(* IEC 61131-3 sources: llm-plc-st-eval/data/processed/gpt-4o/B4/zero_shot, 3 files *)

(* ---- ejec_1.st ---- *)
FUNCTION_BLOCK FB_Giro
VAR_INPUT
    btnFwd : BOOL;   // Botón para giro en sentido horario
    btnRev : BOOL;   // Botón para giro en sentido antihorario
    btnParo : BOOL;  // Botón de paro
END_VAR

VAR_OUTPUT
    fwd : BOOL;      // Salida para giro en sentido horario
    rev : BOOL;      // Salida para giro en sentido antihorario
END_VAR

VAR
    estado : INT;    // Estado actual del motor
END_VAR

// Estados posibles
// 0: Parado
// 1: Girando en sentido horario
// 2: Girando en sentido antihorario

// Lógica de control
IF btnParo THEN
    // Si se presiona el botón de paro, el motor se detiene
    estado := 0;
ELSIF btnFwd AND (estado = 0) THEN
    // Si se presiona el botón de giro horario y el motor está parado
    estado := 1;
ELSIF btnRev AND (estado = 0) THEN
    // Si se presiona el botón de giro antihorario y el motor está parado
    estado := 2;
END_IF

// Actualización de salidas según el estado
CASE estado OF
    0: // Parado
        fwd := FALSE;
        rev := FALSE;
    1: // Girando en sentido horario
        fwd := TRUE;
        rev := FALSE;
    2: // Girando en sentido antihorario
        fwd := FALSE;
        rev := TRUE;
END_CASE

END_FUNCTION_BLOCK

(* ---- ejec_2.st ---- *)
FUNCTION_BLOCK FB_Giro
VAR_INPUT
    btnFwd : BOOL;    // Botón para giro en sentido horario
    btnRev : BOOL;    // Botón para giro en sentido antihorario
    btnParo : BOOL;   // Botón de paro
END_VAR

VAR_OUTPUT
    fwd : BOOL := FALSE;  // Salida para giro en sentido horario
    rev : BOOL := FALSE;  // Salida para giro en sentido antihorario
END_VAR

VAR
    estado : INT := 0;    // Estado del motor: 0 = Parado, 1 = Horario, 2 = Antihorario
END_VAR

// Lógica de control del motor
IF btnParo THEN
    // Si se presiona el botón de paro, detener el motor
    fwd := FALSE;
    rev := FALSE;
    estado := 0;
ELSIF btnFwd AND (estado = 0) THEN
    // Si se presiona el botón de giro horario y el motor está parado
    fwd := TRUE;
    rev := FALSE;
    estado := 1;
ELSIF btnRev AND (estado = 0) THEN
    // Si se presiona el botón de giro antihorario y el motor está parado
    fwd := FALSE;
    rev := TRUE;
    estado := 2;
END_IF
END_FUNCTION_BLOCK

(* ---- ejec_3.st ---- *)
FUNCTION_BLOCK FB_Giro
VAR_INPUT
    btnFwd : BOOL;    // Botón para giro en sentido horario
    btnRev : BOOL;    // Botón para giro en sentido antihorario
    btnParo : BOOL;   // Botón para parar el motor
END_VAR

VAR_OUTPUT
    fwd : BOOL;       // Salida para giro en sentido horario
    rev : BOOL;       // Salida para giro en sentido antihorario
END_VAR

VAR
    estado : INT;     // Estado actual del motor: 0 = Parado, 1 = Horario, -1 = Antihorario
END_VAR

// Inicialización
estado := 0;
fwd := FALSE;
rev := FALSE;

// Lógica de control
IF btnParo THEN
    // Si se presiona el botón de paro, detener el motor
    estado := 0;
    fwd := FALSE;
    rev := FALSE;
ELSIF btnFwd AND (estado = 0) THEN
    // Si se presiona el botón de avance y el motor está parado, girar en sentido horario
    estado := 1;
    fwd := TRUE;
    rev := FALSE;
ELSIF btnRev AND (estado = 0) THEN
    // Si se presiona el botón de retroceso y el motor está parado, girar en sentido antihorario
    estado := -1;
    fwd := FALSE;
    rev := TRUE;
END_IF;
